Fanuc KAREL source: ka00002.KL

PROGRAM KA00002
%STACKSIZE=65535
%PRIORITY=65535
%NOLOCKGROUP
VAR
SRC : INTEGER
DST : REAL
BEGIN
SRC=2
DST=SRC
END KA00002
